//{attribute 'qualified_only'}
VAR_GLOBAL CONSTANT
	ProgramVersion: 			STRING	:=	'V0.1.0.0';			(*	Product . Major . Revision . Build	*)
(*
V0.1.0.0 	- Start version menager.
				- ...

*)	
END_VAR

(* stored: Version 1.1.0.1, ProductVersion 3.1.4024.13
   GVL VersionDescription: Id {3f949215-210a-40c2-bd83-6de6a313f701} *)
